(* PLC project c.project, CODESYS CODESYS V3.5 SP17 Patch 3 *)
(* stored: creationDateTime 2026-10-19T00:00:00, modificationDateTime 2026-10-19T00:00:00 *)

FUNCTION_BLOCK FB_ProbeFbdEno
VAR_INPUT
    xEn : BOOL;
    iSp : INT;
END_VAR
VAR_OUTPUT
    iOut : INT;
    xMoved : BOOL;
END_VAR

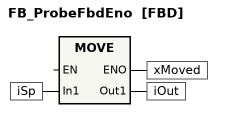
(* FBD diagram, written out as Structured Text *)
xMoved := TRUE;
iOut := iSp;
END_FUNCTION_BLOCK
